SUBAPPLICATION Uebung_094b3d_AX (* Wie Uebung_094b3c_AX (K=2 aktiviert zwei Optionsgruppen NACHEINANDER), aber mit dem neuen generischen T-Stueck Option::splitting::AOption_T_2 statt eines speziellen Weiterleitungs-Plugs auf der Optionsgruppe selbst: OptionalGroup_001 und OptionalGroup_001b sind beide die einfache, unveraenderte Variante (nur ein OPTION-Socket) - das T-Stueck sitzt extern zwischen DEMUX und den beiden Gruppen und kann genauso an eine dritte Gruppe (oder ein weiteres T-Stueck) weitergereicht werden. *)
  (* Standard: 61499-2; Description: Copyright (c) 2026 Meisterschulen am Ostbahnhof This program and the accompanying materials are made available under the terms of the Eclipse Public License 2.0 which is available at https://www.eclipse.org/legal/epl-2.0/ SPDX-License-Identifier: EPL-2.0 *)
  (* Version 1.0, 2026-10-14, Franz Höpfinger, Meisterschulen am Ostbahnhof, initial implementation - zeigt das neue, kaskadierbare T-Stueck AOption_T_2 (Option::splitting) als generische Alternative zum Ad-hoc-PLUG1-Muster aus OptionalGroup_001a/Uebung_094b3c_AX: AOption_AUI_DEMUX_3.OUT2 -> AOption_T_2.IN -> zuerst OUT2 (OptionalGroup_001), danach erst OUT1 (OptionalGroup_001b) - sequenziell nacheinander, nicht gleichzeitig. *)
  PACKAGE Uebungen;
  IMPORT Uebungen::const::UT::DefaultPool::InputNumber_I1;
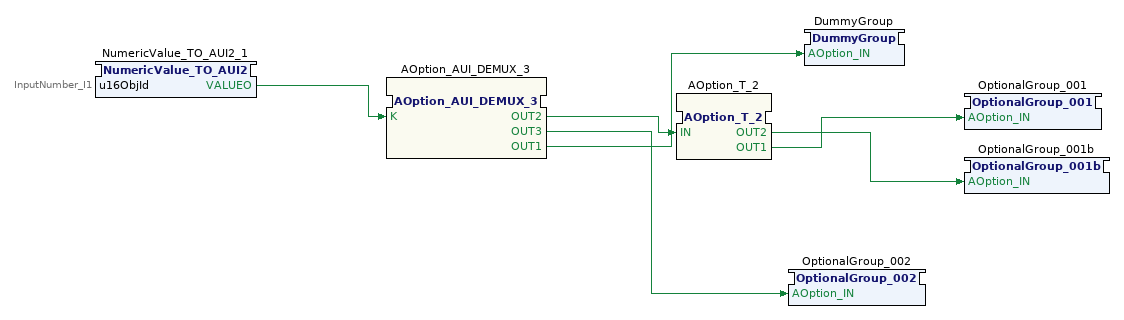
  FBS
    AOption_AUI_DEMUX_3 : Option::selection::AOption_AUI_DEMUX_3;
    AOption_T_2 : Option::splitting::AOption_T_2;
  END_FBS
  SUBAPPS
    NumericValue_TO_AUI2_1 : MyLib::sys::NumericValue_TO_AUI2(u16ObjId := InputNumber_I1);
    OptionalGroup_001 : MyLib_AX_Option::sys::OptionalGroup_001;
    OptionalGroup_001b : MyLib_AX_Option::sys::OptionalGroup_001b;
    OptionalGroup_002 : MyLib_AX_Option::sys::OptionalGroup_002;
    DummyGroup : MyLib_AX_Option::sys::DummyGroup;
  END_SUBAPPS
  ADAPTER_CONNECTIONS
    NumericValue_TO_AUI2_1.VALUEO TO AOption_AUI_DEMUX_3.K;
    AOption_AUI_DEMUX_3.OUT2 TO AOption_T_2.IN;
    AOption_T_2.OUT2 TO OptionalGroup_001b.AOption_IN;
    AOption_AUI_DEMUX_3.OUT3 TO OptionalGroup_002.AOption_IN;
    AOption_AUI_DEMUX_3.OUT1 TO DummyGroup.AOption_IN;
    AOption_T_2.OUT1 TO OptionalGroup_001.AOption_IN;
  END_CONNECTIONS
END_SUBAPPLICATION
